// TIA Portal V21 export
// export: Created 2026-11-02T03:26:15.7867481Z, ExportSetting WithDefaults, DisplayName Totally Integrated Automation Portal, DisplayVersion V21 Update 3, DisplayName TIA Portal Test Suite Advanced, DisplayVersion V21 Update 1, DisplayName SINAMICS Startdrive Advanced, DisplayVersion V21 Update 1, DisplayName SINAMICS Startdrive G130, G150, S120, S150, G200, G210, G210C, G210X, G220, S200, S210, S220, Innomotics MVD, DisplayVersion V21 Update 1, DisplayName SINAMICS Startdrive G110M, G120, G120C, G120D, G120P, G115D, DisplayVersion V21 Update 1, DisplayName STEP 7 Professional, DisplayVersion V21 Update 3, DisplayName STEP 7 Safety, DisplayVersion V21, DisplayName Tech WebApplication, DisplayVersion V21, DisplayName WinCC Basic/Comfort/Advanced, DisplayVersion V21 Update 3, DisplayName WinCC Professional, DisplayVersion V21 Update 3, DisplayName WinCC Unified, DisplayVersion V21 Update 3
DATA_BLOCK "Tgp_InstanceEffect_DB"   // DB2
VERSION : 0.1
// stored: AutoNumber true, DBAccessibleFromOPCUA true, DBAccessibleFromWebserver true, InstanceOfName Tgp_InstanceEffect, InstanceOfType FB
"Tgp_InstanceEffect"
   // VAR_INPUT
   //    Enable : Bool;
   // END_VAR
   // VAR_OUTPUT
   //    Active : Bool;
   // END_VAR
   // VAR
   //    RetainedMarker : Int := 42;
   //    Child { S7_SetPoint := 'True'} : "Tgp_TemplateFB_LAD";
   // END_VAR
BEGIN
END_DATA_BLOCK
